(* PLC project g_estop_reset, Anonymous Benchmark Suite 1.0 *)
(* stored: creationDateTime 2026-08-28T00:00:00 *)

PROGRAM g_estop_reset
  VAR_INPUT
    EStop : BOOL;
    Reset : BOOL;
    Start : BOOL;
  END_VAR
  VAR_OUTPUT
    ResetEdge : BOOL;
    Safe : BOOL;
    Run : BOOL;
    Reset_prev : BOOL;
  END_VAR

(* LD diagram, written out as Structured Text *)
ResetEdge := Reset_prev AND NOT Reset;
Safe := (Safe OR ResetEdge) AND NOT EStop;
Run := Safe AND Start AND NOT EStop;
Reset_prev := Reset;
END_PROGRAM

CONFIGURATION Config0
  RESOURCE Res0 ON PLC
    TASK tcyclic(INTERVAL := T#10ms, PRIORITY := 0);
    PROGRAM inst0 WITH tcyclic : g_estop_reset;
  END_RESOURCE
END_CONFIGURATION
